{attribute 'qualified_only'}
VAR_GLOBAL
	
coffees			: coffee;
teas			: tea;

END_VAR

(* stored: Version 1.1.0.1
   GVL gvl: Id {441aa837-a1ce-4b73-89c3-75f06569f355} *)
